Fanuc KAREL source: KT00027.KL

PROGRAM KT00027
%NOLOCKGROUP
VAR
  H1: ARRAY[2] OF SHORT
  R2: REAL
  OUT: INTEGER
BEGIN
  H1[1] = 2
    R2 = 3.0
  OUT = H1[1] + R2
END KT00027
